(* IEC 61131-3 sources: PLC-Static-Analysis/modules/plc-rules/src/test/resources/PLCA-L004, 2 files *)

(* ---- compliant.st ---- *)
FUNCTION F_Next : INT
F_Next := 1;
END_FUNCTION

PROGRAM P_L004ok
VAR
    n : INT;
    m : INT;
    r : REAL;
    b : BOOL;
    c : BOOL;
    q : BOOL;
    sName : STRING(10);
END_VAR
VAR CONSTANT
    cOn : BOOL := TRUE;
END_VAR
IF n = 1 OR n = 2 THEN
    q := TRUE;
END_IF
q := r <> r;
q := F_Next() > 10 AND F_Next() < 5;
q := cOn AND NOT cOn;
q := n > 10 AND m < 5;
q := sName = 'A' OR sName = 'a';
END_PROGRAM

(* ---- noncompliant.st ---- *)
PROGRAM P_L004
VAR
    n : INT;
    m : INT;
    r : REAL;
    b : BOOL;
    c : BOOL;
    q : BOOL;
    sName : STRING(10);
END_VAR
IF n = 1 AND n = 2 THEN // PLCA-L004
    q := TRUE;
END_IF
q := n > 10 AND n < 5; // PLCA-L004
q := b AND c AND NOT b; // PLCA-L004
WHILE n <> n DO // PLCA-L004
    n := n + 1;
END_WHILE
q := (n > 10 AND m > 3) AND (n < 0 OR n < 5); // PLCA-L004
q := sName = 'A' AND sName = 'a'; // PLCA-L004 (texts compare case-sensitively)
END_PROGRAM
